Fanuc KAREL source: kb00135.KL

-- PROVISIONAL review KL for V1013-1; original PC SHA256 6d1e1a33264cec964a846aa6f2be7d6f74d9ff782cc8f9add28bd7db33bf716f
-- Incomplete behavior may be omitted. Consult companion uncertainty JSON. Do not deploy.
PROGRAM KB00135
%NOLOCKGROUP
BEGIN
  -- UNRESOLVED_PC offsets 5-12; opcodes 9D,23
  -- UNRESOLVED_PC offsets 17-26; opcodes 3F,75
  -- UNRESOLVED_PC offsets 31-38; opcodes 9D,23
  -- UNRESOLVED_PC offsets 43-50; opcodes 9D,23
  -- UNRESOLVED_PC offsets 55-85; opcodes 27,22,22,2A,22,22,31
  -- UNRESOLVED_PC offsets 90-94; opcodes 7F
END KB00135
